(* IEC 61131-3 sources: trust-platform/examples/plant_demo/src, 4 files *)

(* ---- types.st ---- *)
TYPE
    PumpState : (Idle := 0, Starting := 1, Running := 2, Fault := 3);

    PumpCommand :
    STRUCT
        Enable : BOOL;
        TargetSpeed : REAL;
    END_STRUCT;

    PumpStatus :
    STRUCT
        Running : BOOL;
        State : PumpState;
        ActualSpeed : REAL;
        Alarm : UDINT;
    END_STRUCT;
END_TYPE

(* ---- fb_pump.st ---- *)
FUNCTION_BLOCK PumpController
VAR_INPUT
    Command : PumpCommand;
END_VAR
VAR_OUTPUT
    Status : PumpStatus;
END_VAR
VAR
    RampTimer : TON;
    Ramp : REAL;
END_VAR
VAR CONSTANT
    RampTime : TIME := T#1s;
END_VAR

Status.Running := FALSE;
Status.Alarm := 0;

IF NOT Command.Enable THEN
    Status.State := PumpState#Idle;
    Status.ActualSpeed := 0.0;
    Ramp := 0.0;
    RampTimer(IN := FALSE);
ELSE
    CASE Status.State OF
        PumpState#Idle:
            Status.State := PumpState#Starting;
            RampTimer(IN := TRUE, PT := RampTime);
        PumpState#Starting:
            RampTimer(IN := TRUE, PT := RampTime);
            IF RampTimer.Q THEN
                Status.State := PumpState#Running;
            ELSE
                Ramp := Ramp + 0.2;
            END_IF
        PumpState#Running:
            Status.Running := TRUE;
            Ramp := Command.TargetSpeed;
        PumpState#Fault:
            Status.Running := FALSE;
            Status.Alarm := 16#BEEF;
    END_CASE
END_IF

Status.ActualSpeed := Ramp;
END_FUNCTION_BLOCK

(* ---- config.st ---- *)
CONFIGURATION PlantDemo
TASK Fast (INTERVAL := T#100ms, PRIORITY := 1);
PROGRAM P1 WITH Fast : PlantProgram;
VAR_CONFIG
    P1.StartCmd AT %IX0.0 : BOOL;
    P1.SpeedRaw AT %IW0 : INT;
    P1.HaltReq AT %QX0.0 : BOOL;
END_VAR
END_CONFIGURATION

(* ---- program.st ---- *)
PROGRAM PlantProgram
VAR
    Pump : PumpController;
    Cmd : PumpCommand;
    Status : PumpStatus;
    StartCmd : BOOL;
    SpeedRaw : INT;
    SpeedSet : REAL;
    HaltReq : BOOL;
END_VAR

Cmd.Enable := StartCmd AND NOT HaltReq;
SpeedSet := INT_TO_REAL(SpeedRaw);
Cmd.TargetSpeed := SpeedSet;

Pump(Command := Cmd);
Status := Pump.Status;
HaltReq := FALSE;
IF Status.State = PumpState#Fault THEN
    HaltReq := TRUE;
END_IF
END_PROGRAM
